(* IEC 61131-3 sources: codesys-to-s7/tests/corpus/C2S7-SEM-TIMER-Q/pos, 1 file *)

(* ---- input.st ---- *)
FUNCTION_BLOCK FB_Case
VAR
    tPulse : TON;
END_VAR
tPulse(IN := NOT tPulse.Q, PT := T#1S);
END_FUNCTION_BLOCK
